(* PLC project PR_MultiPosShuttle_Soft2.0 1_workflow_268c4d_PLC, SiemensToBackhoff Siemens TIA Portal → Beckhoff TwinCAT PLCopen Converter 2.2 *)
(* stored: creationDateTime 2026-10-12T09:25:10.453821, modificationDateTime 2026-10-12T09:25:10.453821 *)

FUNCTION_BLOCK PR_MultiPosShuttle_Soft2.0 1_workflow_268c4d
VAR_INPUT
	iAutoRunning : BOOL;
	iFaultReset : BOOL;
	iGantry2Safe : BOOL;
	iGantry_2Safe : BOOL;
	iHIPOTTesSafe : BOOL;
	iHIPOTTestOver : BOOL;
	iHipotTestSafe : BOOL;
	iInfeedGantrySafe : BOOL;
	iOTS_Frm_Gantry : BOOL;
	iPartPresent : BOOL;
	iPartPrsent : BOOL;
	iRTR_Frm_Gantry2 : BOOL;
	iReset_fault : BOOL;
	iShuttleAtGantry2Pos : BOOL;
	iShuttleAtGantry_2Pos : BOOL;
	iShuttleAtHIPOTPos : BOOL;
	iShuttleAtHIPOTTestPos : BOOL;
	iShuttleAtPartLoadPos : BOOL;
	iSstMode : BOOL;
	iSstPB : BOOL;
END_VAR
VAR_OUTPUT
	qError : ARRAY[0..10] OF BOOL;
	qHiPotTestStartCmd : BOOL;
	qMessage : ARRAY[0..10] OF BOOL;
	qRTR_To_InfeedGantry : BOOL;
	qShuttleGantry_2PosCmd : BOOL;
	qShuttleHIPOTTestPosCmd : BOOL;
	qStateNo : INT;
	qShuttleReceivePosCmd : BOOL;
END_VAR
VAR
	c10_ChkRecCond_T1 : BOOL;
	c10_ChkRecCond_T2 : BOOL;
	c10_ChkRecCond_T3 : BOOL;
	c10_ChkRecCond_T4 : BOOL;
	c10_ChkRecCond_T5 : BOOL;
	c150_ChkOprnSts_T1 : BOOL;
	c150_ChkOprnSts_T2 : BOOL;
	c30_ChkPartPrsnt_T1 : BOOL;
	c30_ChkPartPrsnt_T2 : BOOL;
	s100_WtHipotTestOver : BOOL;
	s100_WtHipotTestOver_T1 : BOOL;
	s10_ChkRecCond : BOOL;
	s10_ChkRecCond_T1 : BOOL;
	s10_ChkRecCond_T2 : BOOL;
	s10_ChkRecCond_T3 : BOOL;
	s10_ChkRecCond_T4 : BOOL;
	s10_ChkRecCond_T5 : BOOL;
	s110_WtGantry2Safe : BOOL;
	s110_WtGantry2Safe_T1 : BOOL;
	s120_WtShtlGantry2Pos : BOOL;
	s120_WtShtlGantry2Pos_T1 : BOOL;
	s130_WtRTRFrmGantry2 : BOOL;
	s130_WtRTRFrmGantry2_T1 : BOOL;
	s140_WtPartAbsntGantry2Safe : BOOL;
	s140_WtPartAbsntGantry2Safe_T1 : BOOL;
	s150_ChkOprnSts : BOOL;
	s150_ChkOprnSts_T1 : BOOL;
	s150_ChkOprnSts_T2 : BOOL;
	s1_WtResetRel : BOOL;
	s1_WtResetRel_T1 : BOOL;
	s20_WtFaultReset : BOOL;
	s20_WtFaultReset_T1 : BOOL;
	s30_ChkPartPrsnt : BOOL;
	s30_ChkPartPrsnt_T1 : BOOL;
	s30_ChkPartPrsnt_T2 : BOOL;
	s40_WtAllSysSafe : BOOL;
	s40_WtAllSysSafe_T1 : BOOL;
	s50_WtShtlPartRcvPos : BOOL;
	s50_WtShtlPartRcvPos_T1 : BOOL;
	s60_WtOTSFrmGantry : BOOL;
	s60_WtOTSFrmGantry_T1 : BOOL;
	s70_WtPartPlcdGantrySafe : BOOL;
	s70_WtPartPlcdGantrySafe_T1 : BOOL;
	s80_WtHIPOTSafe : BOOL;
	s80_WtHIPOTSafe_T1 : BOOL;
	s90_WtShtlHIPOTPos : BOOL;
	s90_WtShtlHIPOTPos_T1 : BOOL;
	sHIPOTOprnOver : BOOL;
	sHipotTestInProgress : BOOL;
	sPickInProgress : BOOL;
	sPlaceInProgress : BOOL;
	sSst : BOOL;
	sSstPulse : BOOL;
	sSstRise : R_TRIG;
	sStWtResetRel : BOOL;
	sStWtResetRel_T1 : BOOL;
END_VAR
VAR_TEMP
	tOne : BOOL;
END_VAR
  VAR  (* added by the conversion: wires and edge detectors of the diagram *)
    _w24 : BOOL;
    _w26 : BOOL;
    _w39 : BOOL;
    _w41 : BOOL;
    _w42 : BOOL;
    _w99 : BOOL;
    _w102 : BOOL;
    _w103 : BOOL;
    _w104 : BOOL;
    _w105 : BOOL;
    _w106 : BOOL;
    _w107 : BOOL;
    _w120 : BOOL;
    _w122 : BOOL;
    _w123 : BOOL;
    _w151 : BOOL;
    _w154 : BOOL;
    _w155 : BOOL;
    _w156 : BOOL;
    _w171 : BOOL;
    _w173 : BOOL;
    _w174 : BOOL;
    _w187 : BOOL;
    _w189 : BOOL;
    _w190 : BOOL;
    _w207 : BOOL;
    _w209 : BOOL;
    _w210 : BOOL;
    _w228 : BOOL;
    _w231 : BOOL;
    _w232 : BOOL;
    _w251 : BOOL;
    _w254 : BOOL;
    _w255 : BOOL;
    _w268 : BOOL;
    _w270 : BOOL;
    _w271 : BOOL;
    _w289 : BOOL;
    _w292 : BOOL;
    _w293 : BOOL;
    _w312 : BOOL;
    _w315 : BOOL;
    _w316 : BOOL;
    _w333 : BOOL;
    _w335 : BOOL;
    _w336 : BOOL;
    _w353 : BOOL;
    _w355 : BOOL;
    _w356 : BOOL;
    _w370 : BOOL;
    _w373 : BOOL;
    _w374 : BOOL;
    _w404 : BOOL;
    _w406 : BOOL;
    _w407 : BOOL;
    _w408 : BOOL;
  END_VAR

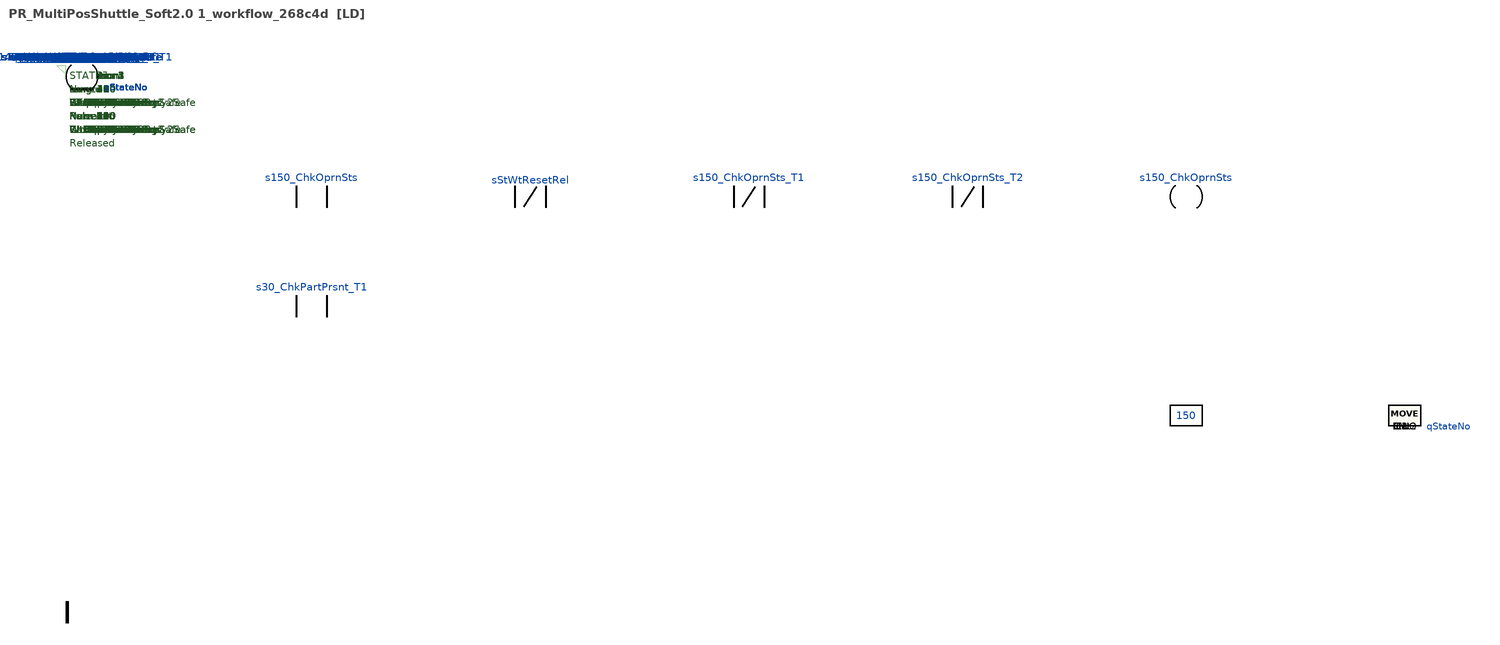
(* LD diagram, written out as Structured Text *)
(* Network 1 *)
(* Create Single Step Pulse bit *)
(* Create Single Step bit *)
(* Transition for STATE Num:0 Reset Released *)
(* STATE Num:0 Reset Released *)
(* Transition for STATE Num:1 WtResetRel *)
(* STATE Num:1 WtResetRel *)
(* Condition1 for STATE Num:10 ChkRecCond *)
(* Condition2 for STATE Num:10 ChkRecCond *)
(* Condition3 for STATE Num:10 ChkRecCond *)
(* Condition4 for STATE Num:10 ChkRecCond *)
(* Condition5 for STATE Num:10 ChkRecCond *)
(* Transition for STATE Num:10 ChkRecCond *)
(* STATE Num:10 ChkRecCond *)
(* Transition for STATE Num:20 WtFaultReset *)
(* STATE Num:20 WtFaultReset *)
(* Actions for STATE Num:20 WtFaultReset *)
(* Condition1 for STATE Num:30 ChkPartPrsnt *)
(* Condition2 for STATE Num:30 ChkPartPrsnt *)
(* Transition for STATE Num:30 ChkPartPrsnt *)
(* STATE Num:30 ChkPartPrsnt *)
(* Transition for STATE Num:40 WtAllSysSafe *)
(* STATE Num:40 WtAllSysSafe *)
(* Transition for STATE Num:50 WtShtlPartRcvPos *)
(* STATE Num:50 WtShtlPartRcvPos *)
(* Actions for STATE Num:50 WtShtlPartRcvPos *)
(* Transition for STATE Num:60 WtOTSFrmGantry *)
(* STATE Num:60 WtOTSFrmGantry *)
(* Actions for STATE Num:60 WtOTSFrmGantry *)
(* Transition for STATE Num:70 WtPartPlcdGantrySafe *)
(* STATE Num:70 WtPartPlcdGantrySafe *)
(* Actions for STATE Num:70 WtPartPlcdGantrySafe *)
(* Transition for STATE Num:80 WtHIPOTSafe *)
(* STATE Num:80 WtHIPOTSafe *)
(* Transition for STATE Num:90 WtShtlHIPOTPos *)
(* STATE Num:90 WtShtlHIPOTPos *)
(* Actions for STATE Num:90 WtShtlHIPOTPos *)
(* Transition for STATE Num:100 WtHipotTestOver *)
(* STATE Num:100 WtHipotTestOver *)
(* Actions for STATE Num:100 WtHipotTestOver *)
(* Transition for STATE Num:110 WtGantry2Safe *)
(* STATE Num:110 WtGantry2Safe *)
(* Actions for STATE Num:110 WtGantry2Safe *)
(* Transition for STATE Num:120 WtShtlGantry2Pos *)
(* STATE Num:120 WtShtlGantry2Pos *)
(* Actions for STATE Num:120 WtShtlGantry2Pos *)
(* Transition for STATE Num:130 WtRTRFrmGantry2 *)
(* STATE Num:130 WtRTRFrmGantry2 *)
(* Transition for STATE Num:140 WtPartAbsntGantry2Safe *)
(* STATE Num:140 WtPartAbsntGantry2Safe *)
(* Actions for STATE Num:140 WtPartAbsntGantry2Safe *)
(* Condition1 for STATE Num:150 ChkOprnSts *)
(* Condition2 for STATE Num:150 ChkOprnSts *)
(* Transition for STATE Num:150 ChkOprnSts *)
(* STATE Num:150 ChkOprnSts *)
tOne := tOne OR NOT tOne;
sSstRise(CLK := iSstPB);
sSstPulse := sSstRise.Q;
sSst := iSstMode AND sSstPulse OR NOT iSstMode;
sStWtResetRel_T1 := sStWtResetRel AND iAutoRunning;
_w24 := sStWtResetRel;
_w26 := (_w24 OR NOT iAutoRunning) AND NOT sStWtResetRel_T1;
sStWtResetRel := _w26;
IF _w26 THEN qStateNo := 0; END_IF;
s1_WtResetRel_T1 := s1_WtResetRel AND NOT sStWtResetRel AND sSst AND iAutoRunning;
_w39 := s1_WtResetRel;
_w41 := (_w39 OR sStWtResetRel_T1) AND NOT sStWtResetRel;
_w42 := _w41 AND NOT s1_WtResetRel_T1;
s1_WtResetRel := _w42;
IF _w42 THEN qStateNo := 1; END_IF;
c10_ChkRecCond_T1 := NOT iPartPrsent AND iShuttleAtHIPOTPos OR NOT iPartPresent AND iShuttleAtGantry_2Pos;
c10_ChkRecCond_T2 := sPickInProgress;
c10_ChkRecCond_T3 := sHipotTestInProgress;
c10_ChkRecCond_T4 := sPlaceInProgress;
c10_ChkRecCond_T5 := NOT sPickInProgress AND NOT sHipotTestInProgress AND NOT sPlaceInProgress AND NOT c10_ChkRecCond_T1;
s10_ChkRecCond_T1 := s10_ChkRecCond AND NOT sStWtResetRel AND sSst AND c10_ChkRecCond_T1;
s10_ChkRecCond_T2 := s10_ChkRecCond AND NOT sStWtResetRel AND sSst AND NOT s10_ChkRecCond_T1 AND c10_ChkRecCond_T2;
s10_ChkRecCond_T3 := s10_ChkRecCond AND NOT sStWtResetRel AND sSst AND NOT s10_ChkRecCond_T1 AND NOT s10_ChkRecCond_T1 AND NOT s10_ChkRecCond_T2 AND c10_ChkRecCond_T3;
s10_ChkRecCond_T4 := s10_ChkRecCond AND NOT sStWtResetRel AND sSst AND NOT s10_ChkRecCond_T1 AND NOT s10_ChkRecCond_T1 AND NOT s10_ChkRecCond_T2 AND NOT s10_ChkRecCond_T1 AND NOT s10_ChkRecCond_T2 AND NOT s10_ChkRecCond_T3 AND c10_ChkRecCond_T4;
s10_ChkRecCond_T5 := s10_ChkRecCond AND NOT sStWtResetRel AND sSst AND NOT s10_ChkRecCond_T1 AND NOT s10_ChkRecCond_T1 AND NOT s10_ChkRecCond_T2 AND NOT s10_ChkRecCond_T1 AND NOT s10_ChkRecCond_T2 AND NOT s10_ChkRecCond_T3 AND NOT s10_ChkRecCond_T1 AND NOT s10_ChkRecCond_T2 AND NOT s10_ChkRecCond_T3 AND NOT s10_ChkRecCond_T4 AND c10_ChkRecCond_T5;
_w99 := s10_ChkRecCond;
_w102 := (_w99 OR s1_WtResetRel_T1 OR s20_WtFaultReset_T1) AND NOT sStWtResetRel;
_w103 := _w102 AND NOT s10_ChkRecCond_T1;
_w104 := _w103 AND NOT s10_ChkRecCond_T2;
_w105 := _w104 AND NOT s10_ChkRecCond_T3;
_w106 := _w105 AND NOT s10_ChkRecCond_T4;
_w107 := _w106 AND NOT s10_ChkRecCond_T5;
s10_ChkRecCond := _w107;
IF _w107 THEN qStateNo := 10; END_IF;
s20_WtFaultReset_T1 := s20_WtFaultReset AND NOT sStWtResetRel AND sSst AND iFaultReset;
_w120 := s20_WtFaultReset;
_w122 := (_w120 OR s10_ChkRecCond_T1) AND NOT sStWtResetRel;
_w123 := _w122 AND NOT s20_WtFaultReset_T1;
s20_WtFaultReset := _w123;
IF _w123 THEN qStateNo := 20; END_IF;
qError[1] := s20_WtFaultReset;
c30_ChkPartPrsnt_T1 := iPartPresent;
c30_ChkPartPrsnt_T2 := NOT iPartPresent;
s30_ChkPartPrsnt_T1 := s30_ChkPartPrsnt AND NOT sStWtResetRel AND sSst AND c30_ChkPartPrsnt_T1;
s30_ChkPartPrsnt_T2 := s30_ChkPartPrsnt AND NOT sStWtResetRel AND sSst AND NOT s30_ChkPartPrsnt_T1 AND c30_ChkPartPrsnt_T2;
_w151 := s30_ChkPartPrsnt;
_w154 := (_w151 OR s10_ChkRecCond_T5 OR s140_WtPartAbsntGantry2Safe_T1) AND NOT sStWtResetRel;
_w155 := _w154 AND NOT s30_ChkPartPrsnt_T1;
_w156 := _w155 AND NOT s30_ChkPartPrsnt_T2;
s30_ChkPartPrsnt := _w156;
IF _w156 THEN qStateNo := 30; END_IF;
s40_WtAllSysSafe_T1 := s40_WtAllSysSafe AND NOT sStWtResetRel AND sSst AND iInfeedGantrySafe AND iHipotTestSafe AND iGantry_2Safe;
_w171 := s40_WtAllSysSafe;
_w173 := (_w171 OR s30_ChkPartPrsnt_T2) AND NOT sStWtResetRel;
_w174 := _w173 AND NOT s40_WtAllSysSafe_T1;
s40_WtAllSysSafe := _w174;
IF _w174 THEN qStateNo := 40; END_IF;
s50_WtShtlPartRcvPos_T1 := s50_WtShtlPartRcvPos AND NOT sStWtResetRel AND sSst AND iShuttleAtPartLoadPos;
_w187 := s50_WtShtlPartRcvPos;
_w189 := (_w187 OR s40_WtAllSysSafe_T1) AND NOT sStWtResetRel;
_w190 := _w189 AND NOT s50_WtShtlPartRcvPos_T1;
s50_WtShtlPartRcvPos := _w190;
IF _w190 THEN qStateNo := 50; END_IF;
qShuttleReceivePosCmd := s50_WtShtlPartRcvPos;
s60_WtOTSFrmGantry_T1 := s60_WtOTSFrmGantry AND NOT sStWtResetRel AND sSst AND iOTS_Frm_Gantry;
_w207 := s60_WtOTSFrmGantry;
_w209 := (_w207 OR s50_WtShtlPartRcvPos_T1) AND NOT sStWtResetRel;
_w210 := _w209 AND NOT s60_WtOTSFrmGantry_T1;
s60_WtOTSFrmGantry := _w210;
IF _w210 THEN qStateNo := 60; END_IF;
qRTR_To_InfeedGantry := s60_WtOTSFrmGantry;
s70_WtPartPlcdGantrySafe_T1 := s70_WtPartPlcdGantrySafe AND NOT sStWtResetRel AND sSst AND iPartPresent AND iInfeedGantrySafe;
_w228 := s70_WtPartPlcdGantrySafe;
_w231 := (_w228 OR s10_ChkRecCond_T4 OR s60_WtOTSFrmGantry_T1) AND NOT sStWtResetRel;
_w232 := _w231 AND NOT s70_WtPartPlcdGantrySafe_T1;
s70_WtPartPlcdGantrySafe := _w232;
IF _w232 THEN qStateNo := 70; END_IF;
qMessage[0] := s70_WtPartPlcdGantrySafe;
qMessage[2] := s70_WtPartPlcdGantrySafe;
sPlaceInProgress := s70_WtPartPlcdGantrySafe;
s80_WtHIPOTSafe_T1 := s80_WtHIPOTSafe AND NOT sStWtResetRel AND sSst AND iHipotTestSafe;
_w251 := s80_WtHIPOTSafe;
_w254 := (_w251 OR s150_ChkOprnSts_T1 OR s70_WtPartPlcdGantrySafe_T1) AND NOT sStWtResetRel;
_w255 := _w254 AND NOT s80_WtHIPOTSafe_T1;
s80_WtHIPOTSafe := _w255;
IF _w255 THEN qStateNo := 80; END_IF;
s90_WtShtlHIPOTPos_T1 := s90_WtShtlHIPOTPos AND NOT sStWtResetRel AND sSst AND iShuttleAtHIPOTTestPos;
_w268 := s90_WtShtlHIPOTPos;
_w270 := (_w268 OR s80_WtHIPOTSafe_T1) AND NOT sStWtResetRel;
_w271 := _w270 AND NOT s90_WtShtlHIPOTPos_T1;
s90_WtShtlHIPOTPos := _w271;
IF _w271 THEN qStateNo := 90; END_IF;
qShuttleHIPOTTestPosCmd := s90_WtShtlHIPOTPos;
s100_WtHipotTestOver_T1 := s100_WtHipotTestOver AND NOT sStWtResetRel AND sSst AND iHIPOTTestOver AND iHIPOTTesSafe;
_w289 := s100_WtHipotTestOver;
_w292 := (_w289 OR s10_ChkRecCond_T3 OR s90_WtShtlHIPOTPos_T1) AND NOT sStWtResetRel;
_w293 := _w292 AND NOT s100_WtHipotTestOver_T1;
s100_WtHipotTestOver := _w293;
IF _w293 THEN qStateNo := 100; END_IF;
qMessage[3] := s100_WtHipotTestOver;
sHipotTestInProgress := s100_WtHipotTestOver;
qHiPotTestStartCmd := s100_WtHipotTestOver;
s110_WtGantry2Safe_T1 := s110_WtGantry2Safe AND NOT sStWtResetRel AND sSst AND iGantry_2Safe;
_w312 := s110_WtGantry2Safe;
_w315 := (_w312 OR s150_ChkOprnSts_T2 OR s100_WtHipotTestOver_T1) AND NOT sStWtResetRel;
_w316 := _w315 AND NOT s110_WtGantry2Safe_T1;
s110_WtGantry2Safe := _w316;
IF _w316 THEN qStateNo := 110; END_IF;
qMessage[4] := s110_WtGantry2Safe;
s120_WtShtlGantry2Pos_T1 := s120_WtShtlGantry2Pos AND NOT sStWtResetRel AND sSst AND iShuttleAtGantry2Pos;
_w333 := s120_WtShtlGantry2Pos;
_w335 := (_w333 OR s110_WtGantry2Safe_T1) AND NOT sStWtResetRel;
_w336 := _w335 AND NOT s120_WtShtlGantry2Pos_T1;
s120_WtShtlGantry2Pos := _w336;
IF _w336 THEN qStateNo := 120; END_IF;
qShuttleGantry_2PosCmd := s120_WtShtlGantry2Pos;
s130_WtRTRFrmGantry2_T1 := s130_WtRTRFrmGantry2 AND NOT sStWtResetRel AND sSst AND iRTR_Frm_Gantry2;
_w353 := s130_WtRTRFrmGantry2;
_w355 := (_w353 OR s120_WtShtlGantry2Pos_T1) AND NOT sStWtResetRel;
_w356 := _w355 AND NOT s130_WtRTRFrmGantry2_T1;
s130_WtRTRFrmGantry2 := _w356;
IF _w356 THEN qStateNo := 130; END_IF;
s140_WtPartAbsntGantry2Safe_T1 := s140_WtPartAbsntGantry2Safe AND NOT sStWtResetRel AND sSst AND NOT iPartPresent AND iGantry_2Safe;
_w370 := s140_WtPartAbsntGantry2Safe;
_w373 := (_w370 OR s10_ChkRecCond_T2 OR s130_WtRTRFrmGantry2_T1) AND NOT sStWtResetRel;
_w374 := _w373 AND NOT s140_WtPartAbsntGantry2Safe_T1;
s140_WtPartAbsntGantry2Safe := _w374;
IF _w374 THEN qStateNo := 140; END_IF;
qMessage[1] := s140_WtPartAbsntGantry2Safe;
qMessage[4] := s140_WtPartAbsntGantry2Safe;
sPickInProgress := s140_WtPartAbsntGantry2Safe;
c150_ChkOprnSts_T1 := NOT sHIPOTOprnOver;
c150_ChkOprnSts_T2 := sHIPOTOprnOver;
s150_ChkOprnSts_T1 := s150_ChkOprnSts AND NOT sStWtResetRel AND sSst AND c150_ChkOprnSts_T1;
s150_ChkOprnSts_T2 := s150_ChkOprnSts AND NOT sStWtResetRel AND sSst AND NOT s150_ChkOprnSts_T1 AND c150_ChkOprnSts_T2;
_w404 := s150_ChkOprnSts;
_w406 := (_w404 OR s30_ChkPartPrsnt_T1) AND NOT sStWtResetRel;
_w407 := _w406 AND NOT s150_ChkOprnSts_T1;
_w408 := _w407 AND NOT s150_ChkOprnSts_T2;
s150_ChkOprnSts := _w408;
IF _w408 THEN qStateNo := 150; END_IF;
END_FUNCTION_BLOCK
